(* CODESYS project 485_CAN_4-transparent.project
   Description: This example has the possibility of using three COM Ports. One is used for reading, another for writing and one for both.  The included visualization shows the reading and writing result together with the used parameters. The user can swathe between the read and write port and the two ports, where one is for reading and the other for writing.
   Title: Serial Com with Visualisation

Project tree, tasks and I/O mapping:
  Device : STMicroelectronics-Linux-ARM_64, STMicroelectronics (Shenzhen) R&D Co., Ltd., version 3.5.19.70
    application Application
      libraries: Standard, 3.5.18.0 (System); CAA SerialCom, 3.4.2.0 (CAA Technical Workgroup); CAA Memory, 3.4.1.0 (CAA Technical Workgroup); VisuDialogs, * (System); CAA Types Extern, 3.5.17.0 (CAA Technical Workgroup); CAN API, 1.0.0.3 (3S - Smart Software Solutions GmbH)
      task MAIN_TASK (cyclic, interval 10 ms, priority 0) calls PLC_PRG
      FB/
        function block SERIAL_LINE [ST]: Fb_init, CLOSE
        function block MsgProcessor_EchoST [ST]: ProcessMessage
      Visualisation/
        visualisation SERIAL_LINE_VISU
        visualisation Visualisation
        visualisation CAN_VISU
        visualisation CAN_VIS
      program PLC_PRG [ST]
      Enums/
        data type SERIAL_LINE_MODE
      license
      global variables GVL
      function calculate_angle [ST]
      function calculate_angle_between_line_and_plane [ST]
      function POINT_AXIS [ST]
      data type MFingerData_t
      data type MFingerCmd_t
      data type MFingerInfo_t
      function Angle_trans [ST]
    SoftMotion General Axis Pool
  text list GlobalTextList
  00000000-0000-0000-0000-000000000000|C:\Users\m.lamp\Documents\license.txt
*)

// Device/Application/Enums/SERIAL_LINE_MODE
TYPE SERIAL_LINE_MODE : (SL_READ, SL_WRITE, SL_READWRITE);
END_TYPE

// Device/Application/MFingerData_t
TYPE MFingerData_t :
STRUCT
	 cmd:MFingerCmd_t;
	 info:MFingerInfo_t;
	 dat: ARRAY[1..8] OF BYTE;
END_STRUCT
END_TYPE

// Device/Application/MFingerCmd_t
TYPE MFingerCmd_t :
STRUCT
	 cmd:DWORD:=8;           // 前面的CMD
     Tp:DWORD:=16;        // 目标位置
     Tv:DWORD:=16;        // 目标速度
	 Tc:DWORD:=16;        // 目标电流
    
END_STRUCT
END_TYPE

// Device/Application/MFingerInfo_t
TYPE MFingerInfo_t :
STRUCT
	cmd:DWORD:=8;          // 前面的CMD
    status:DWORD:=8;    // 故障状态 ，0 表示无故障，异常详情：
													// 0 电机正常
													// 1 电机过温告警
													// 2 电机过温保护
													// 3 电机低压保护
													// 4 电机过压保护
													// 5 电机过流保护
													// 6 电机力矩保护
													// 7 电机熔丝位错保护
													// 8 电机堵转保护
													// ...
	
	
    P:DWORD:=12;        // 当前位置，0-4095 对应 0到满行程
    V:DWORD:=12;        // 当前速度，-2048~2047 单位 0.001行程/s
    I:DWORD:=12;        // 当前电流，-2048~2047 单位 0.01A
    F:DWORD:=12;        // 当前位置，0-4095 对应手指压力传感器Adc原始值
END_STRUCT
END_TYPE

// Device/Application/GVL
VAR_GLOBAL
	(* Message count *)
	g_countMsg_ST	: UINT;
	g_countMsg_CFC	: UINT;
	
	(* This data type descripes the configuration of the CANbus Driver *)
	(*g_busConfig		: CAN.DRIVER_CONFIG := (usiNetwork:= 0, uiBaudrate:= 500, ctMessages:= 10);*)
	g_busConfig		: CAN.DRIVER_CONFIG := (usiNetwork:= 0, uiBaudrate:= 1000, ctMessages:= 10);  
	(* Time limit for receiving messages. T#0s:= no time limit *)
	g_tTimeLimit		: TIME := T#5MS;
	
	gCARxMsg	: CAN.RxMessage;
	gCATxMsg	: CAN.RxMessage;
	gMsgOK	: INT:= 0;
	gMsgErr: INT:= 0;
	
	Gtitle: STRING:='CAN 485 TEST';
	gCANRXed:INT:=0;
	
	g485RXed:INT:= 0;
	g485RdBufLen:UINT:= 0;
	g485RdBuf: ARRAY [1..350] OF BYTE;//
	g485RdBuf_TE:ARRAY [1..350] OF BYTE;//
	g485RawData:ARRAY [1..350] OF BYTE;
	g0:ARRAY [1..500] OF BYTE;
	g06:ARRAY [1..6] OF BYTE;
	g_string:ARRAY [1..6] OF BYTE;
	gcalRawData:ARRAY [1..500] OF BYTE;
	
	g_len_rawdata:UINT:=0;
	g_len_caldata:UINT:=0;
	gPoints:ARRAY [1..21,1..3] OF REAL:=[1(63)];//初始值全部为1
	Points22:ARRAY[1..3] OF REAL;
	gFingerAngle: ARRAY [1..15] OF REAL;
	gFingerAngle_last: ARRAY [1..15] OF REAL;
	gFingerAngle_RH:ARRAY [1..15] OF INT;
	gTemp:ARRAY[1..15] OF INT;
	pi:REAL:=3.14159265358979323846;
END_VAR

// Device/Application/PLC_PRG
PROGRAM PLC_PRG
VAR
	(*
	xTwoLines: BOOL;//:= TRUE;
	xTwoLinesOld: BOOL;
	FirstSerialLine: SERIAL_LINE;
	SecondSerialLine: SERIAL_LINE;
	ThirdSerialLine: SERIAL_LINE;
	*)
	com_rs485:SERIAL_LINE;
END_VAR




/// Receive all incoming messages and echos them with CobId +1
VAR	
	(* A CANbus for handling 11bit CobIds *)
	driver11bit		: CAN.CANBus_11bit := (DriverConfig:= g_busConfig);

	(* Handle for an Mask Receiver *)
	hMaskReceiver	: CAN.CAA.HANDLE;
			
	(* Received messages are passed to MessageProcessors. *)
	msgProcessor	: MsgProcessor_EchoST;
	
	(* Defines a mask for the receiver *)
	maskConfig		: CAN.RECEIVER_MASK := (
										dwIdValue:= 0, 
										dwIdMask:= 0, 
										xRTRValue:= FALSE, 
										xRTRMask:= FALSE, 
										x29BitIdValue:= FALSE, 
										x29BitIdMask:= FALSE, 
										xTransmitValue:= FALSE, 
										xTransmitMask:= TRUE, 
										xAlwaysNewest:= FALSE);

END_VAR

VAR
	canAppState: INT := 100;
	dataIdx:BYTE:=0;
	i:INT;
	cnt:INT;
	
	REC_START :BOOL:=FALSE;
	OFFSET_485 :INT;
	COUNT_485BUF:BYTE:=0;
	COUNT_RAWDATA:INT:=0;
	CAL_START:BOOL;
	CAL_FINAL:BOOL;
	point:BYTE:=1;
	axis:BYTE:=1;
	BUFFER_FINAL:BOOL:=FALSE;
	raw_data_len:UINT;
	j:INT:=1;
	k:BYTE:=1;
	can_count:BYTE:=1;
	
	clear_fault:BOOL:=FALSE;
	temp:INT;
	TON_SEND:TON;
	raw_data_start:UINT:=1;
	raw_data_end:UINT:=1;
	len_raw:UINT:=0;
	len_joint:UINT:=0;
	flag_next:BOOL:=FALSE;
	len_buffer:UINT:=350;
	distance_x:REAL;
	distance_y:REAL;
	distance_z:real;
	
	angle_offset_filter:BYTE:=8;
	angle_smooth_filter:BYTE:=70;
	
	DelayTimer: TON;       // 声明TON定时器实例
    StartDelay: BOOL;      // 触发延时开始的信号（例如按钮按下）
    DelayCompleted: BOOL;  // 延时完成的标志位
	
END_VAR

//This is a example where 3 COM Ports can be used, one for reading, one for writing and one for both
//In the visualization the user can choose the mode (one and two Lines)
//By choosing 2 lines, the First and Second serial line is shown
//By choosing 1 line, the Third serial line is shown

//checks if the visualization has changed and one or two lines should be shown
//checks if the user has switched to one or two lines

(*
IF xTwoLines <> xTwoLinesOld THEN
	IF NOT FirstSerialLine.xClosed THEN
		FirstSerialLine.CLOSE();
		RETURN;
	END_IF
	IF NOT SecondSerialLine.xClosed THEN
		SecondSerialLine.CLOSE();
		RETURN;
	END_IF
	IF NOT ThirdSerialLine.xClosed THEN
		ThirdSerialLine.CLOSE();
		RETURN;
	END_IF
	xTwoLinesOld:= xTwoLines;
END_IF

//set the special parameters for the port
// depending on the Port and the bandwidth the values should be adapted
IF xTwoLines THEN
	FirstSerialLine(
		slMode:= SL_READ, //reading port 
		//udiPort:= 6, //Port number
		udiPort:= 2, //Port number
		//udiBaudrate:= 9600, //bandwidth
		udiBaudrate:= 115200, //bandwidth
		//paParity:= COM.PARITY.EVEN, //the parity is optional
		paParity:= COM.PARITY.NONE,
		sbStopBits:= COM.STOPBIT.ONESTOPBIT,
		udiByteSize := 8); //the stopbits are optional );
	SecondSerialLine(
		slMode:= SL_WRITE,  //writing port
		//udiPort:= 1,
		udiPort:= 2, 
		//udiBaudrate:= 9600,
		udiBaudrate:= 115200, //bandwidth
		//paParity:= COM.PARITY.EVEN,
		paParity:= COM.PARITY.NONE,
		sbStopBits:= COM.STOPBIT.ONESTOPBIT,
		udiByteSize := 8);		
ELSE
	ThirdSerialLine(
	*)
	com_rs485(
		slMode:= SL_READWRITE, 
		//udiPort:= 5,
		udiPort:= 2, 
		udiBaudrate:= 921600,
		//paParity:= COM.PARITY.EVEN,
		paParity:= COM.PARITY.NONE,
		sbStopBits:= COM.STOPBIT.ONESTOPBIT,
		udiByteSize := 8);
//END_IF




/// Configure the CAN Driver
driver11bit(DriverConfig:= g_busConfig, eError=> );

/// Configure MessageProcessor
msgProcessor(CANdriver:= driver11bit);

/// Create a Mask Receiver to receive all messages
/// Each call of GetMaskReceiver generates a new Receiver
IF hMaskReceiver = CAN.CAA.gc_hINVALID THEN
	hMaskReceiver:= driver11bit.GetMaskReceiver(Mask:= maskConfig, eError=> );
END_IF
/// Receive messages and hand them over to the MsgProccessor_Echo
driver11bit.ReceiveMessage(hReceiver:= hMaskReceiver, itfMsgProcessor:= msgProcessor, tTimeLimit:= g_tTimeLimit, eError=> );



IF	clear_fault THEN	//清除故障
	
	
	FOR can_count:=1 TO 15 DO
		gCATxMsg.udiCanId:= can_count;
		gCATxMsg.usiDataLength := 1;
		gCATxMsg.abyData[0]:=16#A5;
		driver11bit.SendMessage(Message:= gCATxMsg, eError=> );
	END_FOR

	clear_fault:=FALSE;
END_IF


DelayTimer(IN := StartDelay, PT := T#30S, Q => DelayCompleted, ET =>);

IF 	canAppState = 100 THEN	
	
	IF g485RXed  <> 0 THEN		
		StartDelay:=FALSE;
		
		g485RXed := 0;
	
		MEM.MemMove(ADR(g485RdBuf), ADR(g485RdBuf_TE), g485RdBufLen);
		
		//拼接数据
		IF g485RdBufLen<320 THEN 
			IF g485RdBuf_TE[1] = 16#0D THEN
				MEM.MemMove(ADR(g485RdBuf_TE), ADR(g485RawData),g485RdBufLen);
				// TODO: 从帧头后的三个 ASCII 字符计算有效数据长度 len_raw
        		// 提示：g485RdBuf_TE[2]、[3]、[4] 为字符 '0'~'9'（ASCII 48~57）
        		// 例如 "305" 表示长度为 305 字节
				len_raw:= 0;//计算长度
				len_joint:=len_joint+g485RdBufLen;
			ELSE
				// TODO: 若非帧头，将后续数据拼接到 g485RawData 已有数据之后
        		// 使用 MemMove 将 g485RdBuf_TE 复制到 g485RawData 的合适偏移位置
        		// 偏移量为当前已拼接长度 len_joint
				
				len_joint:=len_joint+g485RdBufLen;
				// TODO: 判断是否已收齐完整帧（帧头 + 长度字节 + 数据 + 帧尾共 len_raw+6 字节）
				IF 0 THEN
					IF	g485RawData[len_joint]=16#0A THEN
						MEM.MemMove(ADR(g485RawData)+4, ADR(gcalRawData),len_joint-4);
						g_len_caldata:=len_joint-4;
						CAL_START:=TRUE;//开始计算
					ELSE
						MEM.MemMove(ADR(g0), ADR(g485RawData), 500);
					END_IF
					
					len_joint:=0;
					len_raw:=0;
				END_IF
			END_IF
		END_IF
		IF g485RdBufLen>320 THEN
			len_joint:=0;
			IF g485RdBuf_TE[1] = 16#0D THEN
				MEM.MemMove(ADR(g485RdBuf_TE), ADR(g485RawData),g485RdBufLen);
				len_raw:=(g485RdBuf_TE[2]-48)*100+(g485RdBuf_TE[3]-48)*10+(g485RdBuf_TE[4]-48)*1;//计算长度
				IF	g485RawData[len_raw+6]=16#0A THEN
						CAL_START:=TRUE;//开始计算
						g_len_caldata:=g485RdBufLen-4;
						MEM.MemMove(ADR(g485RawData)+4, ADR(gcalRawData),g485RdBufLen-4);
					ELSE
						MEM.MemMove(ADR(g0), ADR(g485RawData), 500);
					END_IF
			END_IF
			
		END_IF
		
		(*//计算这一帧数据的长度
		IF	raw_data_start<len_buffer THEN
			len_raw:=(g485RdBuf_TE[raw_data_start+1]-16#30)*100+(g485RdBuf_TE[raw_data_start+2]-48)*10+(g485RdBuf_TE[raw_data_start+3]-48)*1;
			IF	(raw_data_start+len_raw)>len_buffer THEN//如果超过了这一帧数据就吧剩下的先拷贝完
				MEM.MemMove(ADR(g485RdBuf_TE)+raw_data_start+3, ADR(g485RawData), len_buffer-raw_data_start);
				flag_next:=TRUE;
			ELSE
				IF g485RdBuf_TE[raw_data_start+len_raw+4]=16#0A THEN//判断下一个是不是结尾如果是结尾就开始计算
					MEM.MemMove(ADR(g485RdBuf_TE)+raw_data_start+3, ADR(gcalRawData), len_raw+2);
					CAL_START:=TRUE;//开始计算
					g_len_caldata:=len_raw+2;
				END_IF
			END_IF
		ELSE
			raw_data_start:=1;
		END_IF*)
		
	ELSE
		StartDelay:=TRUE;
	END_IF
	canAppState:= 101;
ELSIF 	canAppState = 101 THEN		
		IF gCANRXed <> 0 THEN
			gCANRXed := 0;
			//CHECK gCARxMsg
			IF gCARxMsg.abyData[0] <> 16#AA THEN
				gCATxMsg.udiCanId:= gCARxMsg.udiCanId-16#100;
				gCATxMsg.usiDataLength := 1;
				gCATxMsg.abyData[0]:=16#A5;
				driver11bit.SendMessage(Message:= gCATxMsg, eError=> );
			
			END_IF
			
			
		END_IF
		canAppState:= 100;
END_IF

IF	DelayTimer.Q THEN
	
	gCATxMsg.usiDataLength := 7;
	gCATxMsg.abyData[0]:=16#AA;
	gCATxMsg.abyData[3]:=16#E8;
	gCATxMsg.abyData[4]:=16#09;
	gCATxMsg.abyData[5]:=16#64;
	gCATxMsg.abyData[6]:=16#03;
	gCATxMsg.abyData[7]:=16#00;
	
	FOR can_count:=1 TO 6 DO
		gCATxMsg.udiCanId:= can_count;
		
		gCATxMsg.abyData[1]:=0;
		gCATxMsg.abyData[2]:=0;
		
		IF	can_count = 2 THEN
			gCATxMsg.abyData[1]:=100;//200
			gCATxMsg.abyData[2]:=2;//0
		END_IF
	
			
		driver11bit.SendMessage(Message:= gCATxMsg, eError=> );
	END_FOR
	StartDelay:=FALSE;
END_IF



IF CAL_START  THEN//开始计算
IF gcalRawData[1]=16#2C AND gcalRawData[g_len_caldata]=16#0A THEN//校验第一位是否对齐
	k:=1;
	axis:=1;
	point:=1;
	MEM.MemMove(ADR(g06), ADR(g_string), 6);//字符串赋空值
	FOR j:=2 TO g_len_caldata-1 DO//获取21个点的坐标值
		IF gcalRawData[j] <> 16#2C THEN
			g_string[k]:=gcalRawData[j];
			k:=k+1;
		ELSE
			IF	g_string[1] = 16#2D THEN //负数
				gPoints[point,axis]:=gPoints[point,axis]*(g_string[2]-16#30)+(g_string[4]-16#30)*0.1+(g_string[5]-16#30)*0.01;
				gPoints[point,axis]:=gPoints[point,axis]*-1;
			ELSE
				gPoints[point,axis]:=gPoints[point,axis]*(g_string[1]-16#30)+(g_string[3]-16#30)*0.1+(g_string[4]-16#30)*0.01;
			END_IF
			axis:=axis+1;
			IF axis=4 THEN
				point:=point+1;
				axis:=1;
			END_IF
			IF point = 22 THEN
				point:=1;
			END_IF
			MEM.MemMove(ADR(g06), ADR(g_string), 6);//字符串赋空值
			k:=1;
		END_IF
	END_FOR
	Points22[1]:=(gPoints[1,1]+gPoints[6,1])/2;
	Points22[2]:=(gPoints[1,2]+gPoints[6,2])/2;
	Points22[3]:=(gPoints[1,3]+gPoints[6,3])/2;
	
	
	
	//计算大拇指
	// TODO: 计算拇指根关节角度（使用 calculate_angle_between_line_and_plane）
	// 直线：由点1→点18 定义；平面：由点6、Points22、点3 确定
	gFingerAngle[1]:=0;
	gFingerAngle[2]:=calculate_angle(POINT_AXIS(gPoints,3),POINT_AXIS(gPoints,1),POINT_AXIS(gPoints,3),POINT_AXIS(gPoints,4));
	
	
	//计算食指
	// TODO: 计算食指近端关节角度（使用 calculate_angle）
	// 计算向量 (点7→点6) 与向量 (点7→点8) 的夹角
	gFingerAngle[3]:=0;
	//计算中指
	// TODO: 计算中指近端关节角度（使用 calculate_angle）
	// 计算向量 (点11→点10) 与向量 (点11→点12) 的夹角
	gFingerAngle[4]:=0;
	//计算无名指
	gFingerAngle[5]:=calculate_angle(POINT_AXIS(gPoints,15),POINT_AXIS(gPoints,14),POINT_AXIS(gPoints,15),POINT_AXIS(gPoints,16));
	//计算小拇指
	gFingerAngle[6]:=calculate_angle(POINT_AXIS(gPoints,19),POINT_AXIS(gPoints,18),POINT_AXIS(gPoints,19),POINT_AXIS(gPoints,20));
	//去抖动
	FOR i:=1 TO 6 DO
		IF	i=1 THEN
			IF	ABS(gFingerAngle[i]-gFingerAngle_last[i])<5 THEN
				gFingerAngle[i]:=gFingerAngle_last[i];
			ELSE
				gFingerAngle_last[i]:=gFingerAngle[i];
			END_IF
			
		ELSE
			// TODO: 其他手指关节突变阈值设为 20°
			IF 0 THEN
				gFingerAngle[i]:=gFingerAngle_last[i];
			ELSE
				gFingerAngle_last[i]:=gFingerAngle[i];
			END_IF
		END_IF
		
		
	END_FOR
	//关节映射
	gFingerAngle_RH[1]:=TO_INT((gFingerAngle_RH[1]*angle_smooth_filter+Angle_trans(gFingerAngle[1],78,85,2000,0)*(100-angle_smooth_filter))/100);
		
		
	gFingerAngle_RH[2]:=TO_INT((gFingerAngle_RH[2]*angle_smooth_filter+Angle_trans(gFingerAngle[2],100,170,4095,0)*(100-angle_smooth_filter))/100);
	
	// TODO: 补全食指关节（索引3）的映射与滤波表达式
	// 输入角度范围 50~170°，输出范围 4095~0	
	gFingerAngle_RH[3]:=TO_INT((gFingerAngle_RH[3]*angle_smooth_filter+ 0 /100);
		
	gFingerAngle_RH[4]:=TO_INT((gFingerAngle_RH[4]*angle_smooth_filter+Angle_trans(gFingerAngle[4],50,170,4095,0)*(100-angle_smooth_filter))/100);
		
	gFingerAngle_RH[5]:=TO_INT((gFingerAngle_RH[5]*angle_smooth_filter+Angle_trans(gFingerAngle[5],50,170,4095,0)*(100-angle_smooth_filter))/100);
		
	gFingerAngle_RH[6]:=TO_INT((gFingerAngle_RH[6]*angle_smooth_filter+Angle_trans(gFingerAngle[6],50,170,4095,0)*(100-angle_smooth_filter))/100);
		
	
	CAL_START:=FALSE;
	CAL_FINAL:=TRUE;
	
	MEM.MemMove(ADR(g0), ADR(gcalRawData), 500);
	
ELSE
	CAL_START:=FALSE;
END_IF
END_IF
 
//header         UID             len      cmd     gFingerAngle    gFingerspeed    gFingercurrent   check 
//0xA5      0X00  0X01-0F       0x07      0xaa      0x00 0x00      0x00  0x00         0x00 0x00    0xsum


IF CAL_FINAL THEN//计算完毕通过CAN发送数据
	gCATxMsg.usiDataLength := 7;
	gCATxMsg.abyData[0]:=16#AA;
	gCATxMsg.abyData[3]:=16#E8;
	gCATxMsg.abyData[4]:=16#09;
	gCATxMsg.abyData[5]:=16#64;
	gCATxMsg.abyData[6]:=16#03;
	gCATxMsg.abyData[7]:=16#00;
	
	FOR can_count:=1 TO 6 DO
		gCATxMsg.udiCanId:= can_count;
		temp:=gFingerAngle_RH[can_count];
		// TODO: 限幅保护，确保 temp 在 0~4095 之间
		IF temp>4095 THEN
			temp:=0;
		ELSIF temp <0 THEN
			temp:=0;
		END_IF
		// TODO: 将 temp 拆分为低字节和高字节，存入 gCATxMsg.abyData[1] 和 [2]
    	// 提示：低字节 = temp MOD 256，高字节 = temp / 256
		gCATxMsg.abyData[1]:=0;
		gCATxMsg.abyData[2]:=0;

		gTemp[can_count]:=temp;
		driver11bit.SendMessage(Message:= gCATxMsg, eError=> );
	END_FOR
	CAL_FINAL:=false;	

END_IF

END_PROGRAM

// Device/Application/calculate_angle_between_line_and_plane
FUNCTION calculate_angle_between_line_and_plane : REAL
VAR_INPUT
	A:ARRAY [1..3] OF REAL;
	B:ARRAY [1..3] OF REAL;
	C:ARRAY [1..3] OF REAL;
	D:ARRAY [1..3] OF REAL;
	E:ARRAY [1..3] OF REAL;
END_VAR
VAR
	i:BYTE;
	VEC_AB: ARRAY[1..3] OF REAL;
	VEC_AC: ARRAY[1..3] OF REAL;
	VEC_DE: ARRAY[1..3] OF REAL;
	VEC_N:ARRAY[1..3] OF REAL;
	dot_product:REAL :=0.0;
	magnitude_N:REAL:=0.0;
	magnitude_DE:REAL:=0.0;
	cos_theta:REAL;
	theta_rad:REAL;
	theta_deg:REAL;
END_VAR

//计算向量AB和AC和DE
FOR i:=1 TO 3 DO 
	VEC_AB[i]:=B[i]-A[i];
	VEC_AC[i]:=C[i]-A[i];
	VEC_DE[i]:=E[i]-D[i];
END_FOR

//计算平面ABC的法向量n，它是AB和AC的叉积  
VEC_N[1]:=VEC_AB[2]*VEC_AC[3]-VEC_AB[3]*VEC_AC[2];
VEC_N[2]:=VEC_AB[3]*VEC_AC[1]-VEC_AB[1]*VEC_AC[3];
VEC_N[3]:=VEC_AB[1]*VEC_AC[2]-VEC_AB[2]*VEC_AC[1];

//计算法向量n和向量DE的点积  
FOR i:=1 TO 3 DO 
	dot_product:=dot_product+(VEC_N[i]*VEC_DE[i]);
END_FOR

//计算模长  
FOR i:=1 TO 3 DO 
	magnitude_N:=magnitude_N+(VEC_N[i]*VEC_N[i]);
	magnitude_DE:=magnitude_DE+(VEC_DE[i]*VEC_DE[i]);
END_FOR
magnitude_N:=SQRT(magnitude_N);
magnitude_DE:=SQRT(magnitude_DE);

//计算夹角的余弦值 
cos_theta := dot_product / (magnitude_N * magnitude_DE);
IF cos_theta>1 THEN
	cos_theta:=1;
ELSIF cos_theta<-1 THEN
	cos_theta:=-1;
END_IF
//计算夹角（线段与平面的夹角是法向量与线段向量夹角的补角）
theta_rad:= ACOS(cos_theta); //结果为弧度
theta_deg:=theta_rad*(180/pi);//转换为角度

calculate_angle_between_line_and_plane:=90-theta_deg;//取补角

END_FUNCTION

// Device/Application/calculate_angle
FUNCTION calculate_angle : REAL
VAR_INPUT
	A:ARRAY [1..3] OF REAL;
	B:ARRAY [1..3] OF REAL;
	C:ARRAY [1..3] OF REAL;
	D:ARRAY [1..3] OF REAL;
END_VAR
VAR
	i:BYTE;
	VEC_AB: ARRAY[1..3] OF REAL;
	VEC_CD: ARRAY[1..3] OF REAL;
	dot_product:REAL :=0.0;
	magnitude_AB:REAL:=0.0;
	magnitude_CD:REAL:=0.0;
	magnitude_ABS:REAL:=0.0;
	magnitude_CDS:REAL:=0.0;
	cos_theta:REAL;
	theta_rad:REAL;
END_VAR

//计算向量AB和AC 
FOR i:=1 TO 3 DO 
	VEC_AB[i]:=B[i]-A[i];
	VEC_CD[i]:=D[i]-C[i];
END_FOR

//计算点积  
FOR i:=1 TO 3 DO 
	dot_product:=dot_product+(VEC_AB[i]*VEC_CD[i]);
END_FOR

//计算模 
FOR i:=1 TO 3 DO 
	magnitude_AB:=magnitude_AB+(VEC_AB[i]*VEC_AB[i]);
	magnitude_CD:=magnitude_CD+(VEC_CD[i]*VEC_CD[i]);
END_FOR
magnitude_ABS:=SQRT(magnitude_AB);
magnitude_CDS:=SQRT(magnitude_CD);
//计算夹角的余弦值 
cos_theta:=dot_product / (magnitude_ABS * magnitude_CDS);

//将余弦值转换为角度（弧度转角度）  
theta_rad:= ACOS(cos_theta); //结果为弧度
calculate_angle:=theta_rad*(180/pi);

END_FUNCTION

// Device/Application/POINT_AXIS
FUNCTION POINT_AXIS : ARRAY[1..3] OF REAL
VAR_INPUT
	POINTS:ARRAY[1..21,1..3]OF REAL;
	A:BYTE;
	
END_VAR
VAR
END_VAR

POINT_AXIS[1]:=POINTS[A,1];
POINT_AXIS[2]:=POINTS[A,2];
POINT_AXIS[3]:=POINTS[A,3];

END_FUNCTION

// Device/Application/Angle_trans
FUNCTION Angle_trans : real
VAR_INPUT
	Ang:REAL;
	ia:INT;
	ib:INT;
	oa:INT;
	ob:INT;
	
END_VAR
VAR
	min_:INT;
	max_:INT;
END_VAR

IF	oa>ob THEN
	min_:=ob;
	max_:=oa;
ELSE
	min_:=oa;
	max_:=ob;
END_IF

IF	ia=ib THEN
	Angle_trans:=oa;
	RETURN;
END_IF
Angle_trans:=(Ang-ia)*(ob-oa)/(ib-ia)+oa;
IF Angle_trans> max_ THEN
	Angle_trans:=max_;
ELSIF Angle_trans<min_ THEN
		Angle_trans:=min_;
END_IF

END_FUNCTION

// Device/Application/FB/SERIAL_LINE
FUNCTION_BLOCK SERIAL_LINE
VAR_INPUT
	slMode: SERIAL_LINE_MODE;
	udiPort: UDINT;
	udiBaudrate: UDINT;
	sbStopBits: COM.STOPBIT:= COM.STOPBIT.ONESTOPBIT;
	paParity: COM.PARITY:= COM.PARITY.EVEN;
	//sWriteText: STRING:= 'Hello World! ';
	//sWriteText: STRING:= '$30 $31 Hello World! ';
	//sWriteText: STRING:= '$7E$11$22$33$44$55$7F';
	sWriteText: STRING:= 'HELLOWOLRD12345689';
	sWriteTextT: STRING;
	udiByteSize: UDINT;
END_VAR
VAR_OUTPUT
	sReadText: STRING;
	errError: COM.ERROR;
	xReadSuccess: BOOL;
	xWriteSuccess: BOOL;
	xClosed: BOOL:= TRUE;
END_VAR
VAR
	iState: INT;
	tTimer: TON;
	comOpen: COM.Open; (* Instance of the function block for opening a port *)
	hCom: CAA.HANDLE; (* handle of the port*)
	aParameter: ARRAY [1..7] OF COM.PARAMETER;
	comWrite: COM.Write;	(* Instance of the Write function  block *)
	bWriteBuffer: ARRAY [1..80] OF BYTE; (*Used to write data to the serial port*)
	szWrite: CAA.SIZE;
	comRead: COM.Read; (* Instance of the Read function block *)
	bReadBuffer: ARRAY [1..350] OF BYTE; (*Used to read data from the serial port*)
	szRead: CAA.SIZE;
	comClose: COM.Close; (* Instance of the function block for closing a port *)
END_VAR

CASE iState OF
	
	0:	// The parameter for the COM Ports are set
		aParameter[1].udiParameterId:= COM.CAA_Parameter_Constants.udiPort;
		aParameter[1].udiValue:= udiPort;
		aParameter[2].udiParameterId:= COM.CAA_Parameter_Constants.udiBaudrate;
		aParameter[2].udiValue:= udiBaudrate;		
		aParameter[3].udiParameterId:= COM.CAA_Parameter_Constants.udiStopBits;
		aParameter[3].udiValue:= INT_TO_UDINT(sbStopBits);
		aParameter[4].udiParameterId:= COM.CAA_Parameter_Constants.udiParity;
		aParameter[4].udiValue:= INT_TO_UDINT(paParity);
		aParameter[5].udiParameterId:= COM.CAA_Parameter_Constants.udiTimeout;
		aParameter[5].udiValue:= 0;
		aParameter[6].udiParameterId:= COM.CAA_Parameter_Constants.udiBinary;
		aParameter[6].udiValue:= 0;
		aParameter[7].udiParameterId:= COM.CAA_Parameter_Constants.udiByteSize;
		aParameter[7].udiValue:= udiByteSize;
		
		iState:= 1;
		
	1:	//First the COM Port is opened
		comOpen(xExecute:= TRUE, usiListLength:= SIZEOF(aParameter) / SIZEOF(COM.PARAMETER), pParameterList:= ADR(aParameter), hCom=> hCom);
		xClosed:= FALSE;
		IF comOpen.xDone THEN
			comOpen(xExecute:= FALSE);
			//depending on the mode the state for reading or writing is set
			IF slMode = SL_READ OR slMode = SL_READWRITE THEN
				iState:= 2;
			ELSIF slMode = SL_WRITE THEN
				iState:= 4;
			END_IF
		ELSIF comOpen.xError THEN
			errError:= comOpen.eError;
			comOpen(xExecute:= FALSE);
			iState:= 32767;
		END_IF
		
	2: //The reading process is started
		comRead(xExecute:= TRUE, hCom:= hCom, pBuffer:= ADR(bReadBuffer), szBuffer:= SIZEOF(bReadBuffer));
		IF comRead.xDone THEN
			szRead:= comRead.szSize;
			//check if the Port has send something
			IF szRead > 0 THEN
				//the text from the read buffer is saved in the sReadText variable
				//MEM.MemMove(ADR(bReadBuffer), ADR(sReadText), ANY_TO_UINT(szRead));
				//MEM.MemFill(ADR(sReadText) + ANY_TO_UINT(szRead), 1, 0);
				xReadSuccess:= TRUE;
				
				MEM.MemMove(ADR(bReadBuffer), ADR(g485RdBuf), ANY_TO_UINT(szRead));
				g485RdBufLen := ANY_TO_INT(szRead);
				g485RXed := 1;
			END_IF
			// the flag has to be set to false, that in the next cylce, the read task will start again, by setting it to true
			comRead(xExecute:= FALSE);
			///iState:= 3;
		ELSIF comRead.xError THEN
			errError:= comRead.eError;
			comRead(xExecute:= FALSE);
			////iState:= 32767;
		END_IF
		
	3: //After the reading process is finished, a timer is started for waiting 250 milliseconds
		tTimer(IN:= TRUE, PT:= T#250MS);
		IF tTimer.Q THEN
			tTimer(IN:= FALSE);
			xReadSuccess:= FALSE;
			IF slMode = SL_READWRITE THEN
				iState:= 4;
			ELSE
				iState:= 2;
			END_IF
		END_IF
		
	4: // the writing process is started
		IF NOT comWrite.xExecute THEN
			;
			sWriteTextT := CONCAT(CONCAT('$7E',sWriteText),'$7F');
			//sWriteText := sWriteTextT;
			;
			szWrite:= INT_TO_UDINT(LEN(sWriteTextT));
			//write the string to the buffer for the COM.WRITE Interface
			MEM.MemMove(ADR(sWriteTextT), ADR(bWriteBuffer), ANY_TO_UINT(szWrite));
		END_IF
		comWrite(xExecute:= TRUE, hCom:= hCom, pBuffer:= ADR(bWriteBuffer), szSize:= szWrite);
		IF comWrite.xDone THEN
			// the flag is set to false, that in the next cyle this process is started again, by setting it to true 
			comWrite(xExecute:= FALSE);	
			xWriteSuccess:= TRUE;
			iState:= 5;
		ELSIF comWrite.xError THEN
			errError:= comWrite.eError;
			comWrite(xExecute:= FALSE);	
			iState:= 32767;
		END_IF 
		
	5: //After the writing process is finished, a timer is started for waiting 250 milliseconds
		tTimer(IN:= TRUE, PT:= T#250MS);
		IF tTimer.Q THEN
			tTimer(IN:= FALSE);
			xWriteSuccess:= FALSE;
			IF slMode = SL_READWRITE THEN
				iState:= 2;
			ELSE
				iState:= 4;
			END_IF
		END_IF
		
	6: //Closing the ports
		IF hCom <> 0 THEN
			comClose(xExecute:= TRUE, hCom:= hCom);
			IF comClose.xDone THEN
				comClose(xExecute:= FALSE);
				Fb_Init(FALSE, FALSE);
			ELSIF comClose.xError THEN
				errError:= comClose.eError;
				comClose(xExecute:= FALSE);	
				iState:= 32767;
			END_IF
		ELSE
			Fb_Init(FALSE, FALSE);
		END_IF 

	32767:
		;

END_CASE

METHOD Fb_init : BOOL
VAR_INPUT
	bInitRetains : BOOL;
  	bInCopyCode : BOOL; 
END_VAR
END_METHOD

ACTION CLOSE:
iState:= 6;
THIS^();
END_ACTION

END_FUNCTION_BLOCK

// Device/Application/FB/MsgProcessor_EchoST
/// MsgProcessor_Echo is the implimentation of IMessageProcessor. 
/// MsgProcessor_Echo simply counts all incoming messages and echos them with CobId +1
FUNCTION_BLOCK MsgProcessor_EchoST IMPLEMENTS CAN.IMessageProcessor
VAR_IN_OUT
	CANdriver	: CAN.CANBus_11bit;
END_VAR
VAR_OUTPUT
END_VAR
VAR
	_pCANdriver : POINTER TO CAN.CANBus_11bit;
END_VAR

_pCANdriver := ADR(CANdriver);

METHOD ProcessMessage
VAR_IN_OUT
	(* The messages received by the receiver *)
	Message	: CAN.RxMessage;
END_VAR
VAR
END_VAR
/// Echo incoming messages with CobId +1
IF _pCANdriver <> 0 THEN	
	gCARxMsg := Message;	
	
	(*
	Message.udiCanId:= Message.udiCanID + 1;
	_pCANdriver^.SendMessage(Message:= Message, eError=> );	
	*)
	g_countMsg_ST:= g_countMsg_ST +1;
	gCANRXed := 1;	
END_IF
END_METHOD

END_FUNCTION_BLOCK

// Device/Application/Visualisation/SERIAL_LINE_VISU
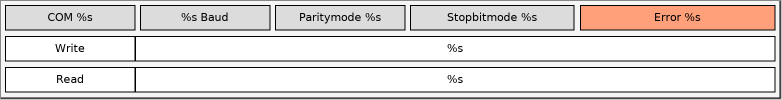
VISUALIZATION SERIAL_LINE_VISU  // 782x100
VAR_IN_OUT
	slInstance: SERIAL_LINE;
END_VAR
    Rectangle (0,0 780x98)
    Rectangle (135,36 640x25), "%s", text variable: slInstance.sWriteText, invisible if: slInstance.slMode = SL_READ
        OnMouseDown: write the text variable via Edit
    Rectangle (5,36 130x25), "Write", colour toggle: slInstance.xWriteSuccess, invisible if: slInstance.slMode = SL_READ
    Rectangle (135,67 640x25), "%s", text variable: slInstance.sReadText, invisible if: slInstance.slMode = SL_WRITE
    Rectangle (5,67 130x25), "Read", colour toggle: slInstance.xReadSuccess, invisible if: slInstance.slMode = SL_WRITE
    Rectangle (5,5 130x25), "COM %s", text variable: slInstance.udiPort
    Rectangle (140,5 130x25), "%s Baud", text variable: slINstance.udiBaudrate
    Rectangle (580,5 195x25), "Error %s", text variable: slInstance.errError
    Rectangle (275,5 130x25), "Paritymode %s", text variable: slInstance.paParity
    Rectangle (410,5 164x25), "Stopbitmode %s", text variable: slInstance.sbStopBits
END_VISUALIZATION

// Device/Application/Visualisation/Visualisation
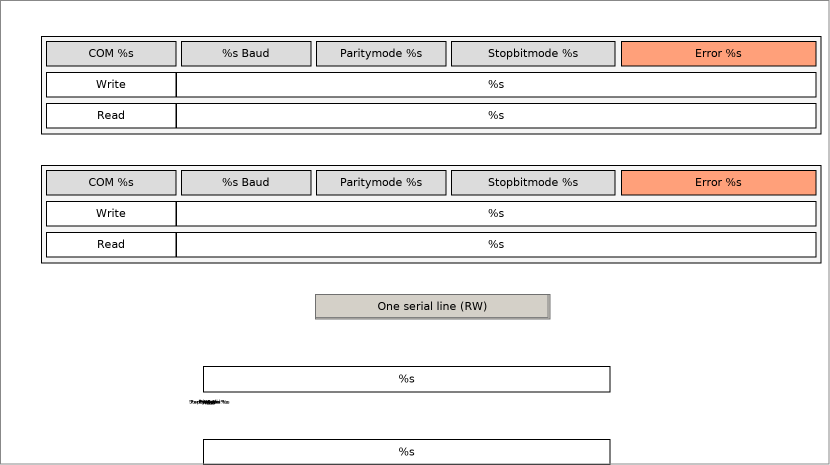
VISUALIZATION Visualisation  // 830x465
AR_IN_OUT
	
END_VAR
    Frame (41,36 787x107), invisible if: NOT PLC_PRG.xTwoLines
        shows SERIAL_LINE_VISU(slInstance := PLC_PRG.FirstSerialLine)
    Frame (41,165 789x109), invisible if: NOT PLC_PRG.xTwoLines
        shows SERIAL_LINE_VISU(slInstance := PLC_PRG.SecondSerialLine)
    Frame (41,36 789x109), invisible if: PLC_PRG.xTwoLines
        shows SERIAL_LINE_VISU(slInstance := PLC_PRG.com_rs485)
    Button (315,294 235x25), "Two serial lines (R / W)", invisible if: PLC_PRG.xTwoLines
        toggle PLC_PRG.xTwoLines
    Button (315,294 235x25), "One serial line (RW)"
    Frame (209,402 1x1)
        shows SERIAL_LINE_VISU()
    Rectangle (203,366 407x26), "%s", text variable: GVL.gCARxMsg.abyData
    Rectangle (203,439 407x26), "%s", text variable: GVL.gCARxMsg.abyData
END_VISUALIZATION

// Device/Application/Visualisation/CAN_VISU
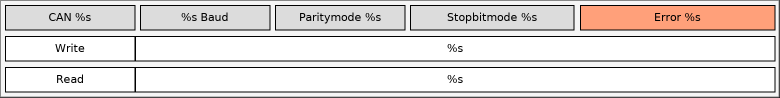
VISUALIZATION CAN_VISU  // 780x98
VAR_IN_OUT
	//slInstance: SERIAL_LINE;
END_VAR
    Rectangle (0,0 780x98)
    Rectangle (135,36 640x25), "%s", text variable: slInstance.sWriteText1, invisible if: slInstance.slMode = SL_READ
        OnMouseDown: write the text variable via Edit
    Rectangle (5,36 130x25), "Write", colour toggle: slInstance.xWriteSuccess, invisible if: slInstance.slMode = SL_READ
    Rectangle (135,67 640x25), "%s", text variable: PLC_PRG.g_CAN_rx_msg
    Rectangle (5,67 130x25), "Read", colour toggle: slInstance.xReadSuccess, invisible if: slInstance.slMode = SL_WRITE
    Rectangle (5,5 130x25), "CAN %s", text variable: slInstance.udiPort
    Rectangle (140,5 130x25), "%s Baud", text variable: slINstance.udiBaudrate
    Rectangle (580,5 195x25), "Error %s", text variable: slInstance.errError
    Rectangle (275,5 130x25), "Paritymode %s", text variable: slInstance.paParity
    Rectangle (410,5 164x25), "Stopbitmode %s", text variable: slInstance.sbStopBits
END_VISUALIZATION

// Device/Application/Visualisation/CAN_VIS
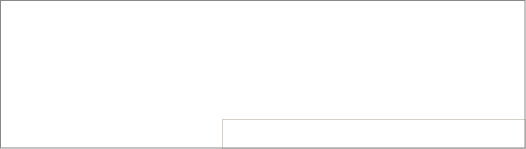
VISUALIZATION CAN_VIS  // 526x149
    Textfield (222,119 304x30)
END_VISUALIZATION
